(* IEC 61131-3 sources: avi-aoi-management/scripts/ai-eval/ngau-nhien/kho/st-ud10-thang-nang-2-tang/khung/src, 2 files *)

(* ---- KhoaDongCo.st ---- *)
FUNCTION_BLOCK KhoaDongCo
VAR_INPUT
    YC_LEN : BOOL;
    YC_XUONG : BOOL;
    CUA_DONG : BOOL;
    DUNG_KHAN : BOOL;
END_VAR
VAR_OUTPUT
    LEN : BOOL;
    XUONG : BOOL;
END_VAR
    (* TODO: cài đặt theo đề bài *)
    LEN := FALSE;
END_FUNCTION_BLOCK

(* ---- ThangNang2Tang.st ---- *)
FUNCTION_BLOCK ThangNang2Tang
VAR_INPUT
    GOI_1 : BOOL;
    GOI_2 : BOOL;
    CT_TANG_1 : BOOL;
    CT_TANG_2 : BOOL;
    CUA_DONG : BOOL;
    DUNG_KHAN : BOOL;
    RESET : BOOL;
    T_DI_CHUYEN : TIME;
END_VAR
VAR_OUTPUT
    LEN : BOOL;
    XUONG : BOOL;
    TRANG_THAI : INT;
    TANG : INT;
    MA_LOI : INT;
END_VAR
    (* TODO: cài đặt theo đề bài *)
    LEN := FALSE;
END_FUNCTION_BLOCK
